Fanuc KAREL source: kt00724.KL

-- PROVISIONAL review KL for V940-1; original PC SHA256 07a3bad19a0185e656c278d5bc96880ab5af1c985db223320df6ad82f49fd379
-- Incomplete behavior may be omitted. Consult companion uncertainty JSON. Do not deploy.
PROGRAM KT00724
%NOLOCKGROUP
VAR
  OUT : BOOLEAN
-- UNRESOLVED_DECL P1 type=000199
-- UNRESOLVED_DECL P2 type=000199
BEGIN
  -- V9_ZERO_TABLE_METADATA_HINT layout=0001; no indexed target words; source/name/runtime held
  -- UNRESOLVED_PC offsets 5-20; opcodes 22,63,23
  -- UNRESOLVED_PC offsets 25-29; opcodes 7F
END KT00724
